(*
SPDX-FileCopyrightText: © 2026 Oleksandr Tiutyk <trofimich@gmail.com>
SPDX-License-Identifier: MIT
License: https://opensource.org/license/mit
*)

(*!
<summary>Checks safe defaults for an unbound TaskRunningSubstate view.</summary>
<description>
Uses unbound local references and checks every observable property without dereferencing a missing target.
</description>
*)

{attribute 'no_explicit_call' := 'do not call this function block directly'}
FUNCTION_BLOCK UnboundTaskRunningSubstateTest EXTENDS TOF_Testing.SingleCycleTest
VAR_STAT
	{attribute 'hide'}
	_ClassName : STRING := __POUNAME();
END_VAR

//! <summary>Reads all flags and verifies the default value for an unbound view.</summary>
METHOD PROTECTED ExecuteTest
VAR
	backingValue : REFERENCE TO TOF_Tasks.TASK_RUNNING_SUBSTATE;
	view : TOF_Tasks.TaskRunningSubstate(taskRunningSubstate := backingValue);
END_VAR
Assert.ThatBool(
	actual := view.ResourceAcquiring,
	message := "Unbound TaskRunningSubstate.ResourceAcquiring must be false"
).IsFalse();
Assert.ThatBool(actual := view.Processing, message := "Unbound TaskRunningSubstate.Processing must be false").IsFalse();
Assert.ThatBool(actual := view.Stopping, message := "Unbound TaskRunningSubstate.Stopping must be false").IsFalse();
Assert.ThatBool(
	actual := view.ResourceReleasing,
	message := "Unbound TaskRunningSubstate.ResourceReleasing must be false"
).IsFalse();
Assert.ThatBool(
	actual := view.Value = TOF_Tasks.TASK_RUNNING_SUBSTATE.RESOURCE_ACQUIRING,
	message := "Unbound Value must default to RESOURCE_ACQUIRING"
).IsTrue();
END_METHOD

//! <summary>Borrows the concrete class name. Callers must not modify the returned storage.</summary>
{attribute 'monitoring' := 'call'}
PROPERTY ClassName : REFERENCE TO STRING
GET
ClassName REF= _ClassName;
END_GET
END_PROPERTY

//! <summary>Borrows the compiler-initialized namespace name. Callers must not modify the returned storage.</summary>
{attribute 'monitoring' := 'call'}
PROPERTY NamespaceName : REFERENCE TO STRING
GET
NamespaceName REF= CurrentNamespace.Name;
END_GET
END_PROPERTY

//! <summary>Reports the complete concrete instance size in bytes.</summary>
{attribute 'monitoring' := 'call'}
PROPERTY SelfSize : ULINT
GET
SelfSize := XSIZEOF(THIS^);
END_GET
END_PROPERTY

END_FUNCTION_BLOCK

(* stored: Version 1.1.0.1
   POU UnboundTaskRunningSubstateTest: Id {8975ddfb-9f1d-44ac-8ece-d30fa7e3dc92}, SpecialFunc None
   Method ExecuteTest: Id {3b3b6c78-a4f0-43be-9f92-630463c99c9e}
   Property ClassName: Id {07e8a124-19c8-4d61-bca0-2f5c0feeee2c}
   Get Get: Id {6ec79182-7732-4500-9f29-e2b8b9a7af6c}
   Property NamespaceName: Id {209ac211-4a3b-4ab3-8858-86c5ca64dec1}
   Get Get: Id {88fad9b4-be2e-4b25-a6c2-8c1dd0404c50}
   Property SelfSize: Id {0f87c90c-f50c-4419-9dbe-28e981369516}
   Get Get: Id {08dd9d92-0eae-4a2d-9b7b-a3863aa1a362} *)
